// Contexte d'un mover dans le séquenceur général (docs/05 § 5.3)
TYPE ST_MoverCtx :
STRUCT
    eState : E_MoverState;
    eWait : E_WaitReason;
    nTable : INT;
    nPC : INT;
    aRetTable : ARRAY[1..GVL_Const.MAX_CALL_DEPTH] OF INT;
    aRetPC : ARRAY[1..GVL_Const.MAX_CALL_DEPTH] OF INT;
    nDepth : USINT;
    nTargetGroup : USINT;
    nTargetOp : USINT;
    nTargetSlot : USINT;
    aOpParam : ARRAY[1..GVL_Const.MAX_PARAMS] OF LREAL;   // paramètres résolus à l'émission de Route
    nStation : USINT;               // station réservée ou occupée, 0 = aucune
    nDest : INT;                    // position planaire de destination
    nPos : INT;                     // position planaire occupée, 0 = entre deux positions
    nReqId : UDINT;
    bRequestPosted : BOOL;
    nRouteRetry : UDINT;
    tWaitStart : LINT;
    fWaitMs : LREAL;
    fMoveMs : LREAL;                // durée du déplacement en cours
    fStillMs : LREAL;               // à l'arrêt dans la fenêtre d'arrivée
    bQualityLock : BOOL;
    bOutOfService : BOOL;
    bImmediate : BOOL;
    bAbsent : BOOL;                 // hors service et absent du plan (D85)
    bStationAborted : BOOL;         // la station de l'opération est passée Aborted (docs/05 § 6.4)
    bToEmptyPark : BOOL;            // en route vers le parcage pour être vidé
    aBadAtArrival : ARRAY[1..GVL_Const.MAX_SLOTS] OF BOOL;     // verdict déjà mauvais à l'arrivée (docs/10 § 9)
    aDefectBad : ARRAY[1..GVL_Const.MAX_SLOTS] OF BOOL;        // mauvaise sur défaut de station (docs/10 § 2)
    aHidden : ARRAY[1..8] OF LREAL; // compteurs de boucle du process général (D93)
    tOpStart : LINT;                // début de l'opération en cours
    fX : LREAL;                     // position actuelle sur le plan
    fY : LREAL;
    fC : LREAL;
    aSlot : ARRAY[1..GVL_Const.MAX_SLOTS] OF ST_Part;
    aVar : ARRAY[1..GVL_Const.MAX_MOVER_VARS] OF LREAL;          // variables de mover (docs/05 § 5.8)
    aVarPos : ARRAY[1..GVL_Const.MAX_MOVER_VARS] OF ST_Position;
    aVarId : ARRAY[1..GVL_Const.MAX_MOVER_VARS] OF UDINT;
END_STRUCT
END_TYPE

(* stored: Version 1.1.0.1, ProductVersion 3.1.4024.12
   DUT ST_MoverCtx: Id {27975211-2829-5c6f-8a6a-eb17e91eab6a} *)
